PROGRAM PRG_IO_Out
VAR
END_VAR

IF GVL_Ctrl.xSim THEN
    // simulation: keep every real output OFF
    GVL_HW.xMaintVent := FALSE;       GVL_HW.xLaserEnable := FALSE;
    GVL_HW.xCW_Trig := FALSE;         GVL_HW.xCW_STO := FALSE;
    GVL_HW.xCW_Job0 := FALSE;  GVL_HW.xCW_Job1 := FALSE;  GVL_HW.xCW_Job2 := FALSE;  GVL_HW.xCW_Job3 := FALSE;
    GVL_HW.xValveInfeed_AS := FALSE;   GVL_HW.xValveInfeed_GS := FALSE;
    GVL_HW.xValveOutfeed_AS := FALSE;  GVL_HW.xValveOutfeed_GS := FALSE;
    GVL_HW.xValveEjector_AS := FALSE;  GVL_HW.xValveEjector_GS := FALSE;
    GVL_HW.xValveClamp_AS := FALSE;    GVL_HW.xValveClamp_GS := FALSE;
    GVL_HW.xValveDiverter_AS := FALSE; GVL_HW.xValveDiverter_GS := FALSE;
    GVL_HW.xValveBlow_AS := FALSE;     GVL_HW.xValveBlow_GS := FALSE;
    GVL_HW.xValveBypass_AS := FALSE;   GVL_HW.xValveBypass_GS := FALSE;
ELSE
    GVL_HW.xMaintVent   := GVL_IO.xVent;
    GVL_HW.xLaserEnable := GVL_IO.xLaserEnable;
    GVL_HW.xCW_Trig     := GVL_IO.xCW_Trig;
    GVL_HW.xCW_STO      := GVL_IO.xCW_STO;
    GVL_HW.xCW_Job0     := (GVL_IO.nCW_Job AND 16#01) <> 0;
    GVL_HW.xCW_Job1     := (GVL_IO.nCW_Job AND 16#02) <> 0;
    GVL_HW.xCW_Job2     := (GVL_IO.nCW_Job AND 16#04) <> 0;
    GVL_HW.xCW_Job3     := (GVL_IO.nCW_Job AND 16#08) <> 0;

    GVL_HW.xValveInfeed_AS   := GVL_IO.stInfeed.xValveWork;    GVL_HW.xValveInfeed_GS   := GVL_IO.stInfeed.xValveHome;
    GVL_HW.xValveOutfeed_AS  := GVL_IO.stOutfeed.xValveWork;   GVL_HW.xValveOutfeed_GS  := GVL_IO.stOutfeed.xValveHome;
    GVL_HW.xValveEjector_AS  := GVL_IO.stEjector.xValveWork;   GVL_HW.xValveEjector_GS  := GVL_IO.stEjector.xValveHome;
    GVL_HW.xValveClamp_AS    := GVL_IO.stClamp.xValveWork;     GVL_HW.xValveClamp_GS    := GVL_IO.stClamp.xValveHome;
    GVL_HW.xValveDiverter_AS := GVL_IO.stDiverter.xValveWork;  GVL_HW.xValveDiverter_GS := GVL_IO.stDiverter.xValveHome;
    GVL_HW.xValveBlow_AS     := GVL_IO.xBlowAS;                GVL_HW.xValveBlow_GS     := GVL_IO.xBlowGS;
    GVL_HW.xValveBypass_AS   := GVL_IO.xBypassAS;              GVL_HW.xValveBypass_GS   := GVL_IO.xBypassGS;
END_IF

END_PROGRAM

(* stored: Version 1.1.0.1
   POU PRG_IO_Out: Id {6b63ea75-6d2f-497d-b8f1-3b625359e5ab}, SpecialFunc None *)
